// TIA Portal V21 export
// export: Created 2026-10-12T12:46:18.6521538Z, ExportSetting WithDefaults, DisplayName Totally Integrated Automation Portal, DisplayVersion V21, DisplayName STEP 7 Professional, DisplayVersion V21, DisplayName STEP 7 Safety, DisplayVersion V21, DisplayName Tech WebApplication, DisplayVersion V21, DisplayName WinCC Basic/Comfort/Advanced, DisplayVersion V21, DisplayName WinCC Unified, DisplayVersion V21
TagTable "IO"
  IB0 : Byte  (%IB0, HMI_Connection_1, 1 s)
  IB1 : Byte  (%IB1, HMI_Connection_1, 1 s)
  QB0 : Byte  (%QB0, HMI_Connection_1, 1 s)
  QB1 : Byte  (%QB1, HMI_Connection_1, 1 s)
